{attribute 'pack_mode' := '1'}
TYPE ST_ProtectionConfig_Rx :
STRUCT
	BatWarrning			:	REAL;
	BatFault			:	REAL;
	BatRoomTempWarrning	:	REAL;
	BatRoomTempFault	:	REAL;
	BatRoomHumWarrning	:	REAL;
	BatRoomHumFault		:	REAL;
END_STRUCT
END_TYPE

(* stored: Version 1.1.0.1, ProductVersion 3.1.4024.9
   DUT ST_ProtectionConfig_Rx: Id {3ac122dd-5f44-4b2e-89e6-43295a74b0d4} *)
